{attribute 'pack_mode' := '1'}
TYPE ST_ModulePublishData :
STRUCT
 Header : ST_MqttHeader;
 Devices : ARRAY[0..GVL_PARAM.BAT_MODULE_COUNT-1] OF ST_ModulePublish_V1;
END_STRUCT
END_TYPE

(* stored: Version 1.1.0.1, ProductVersion 3.1.4024.15
   DUT ST_ModulePublishData: Id {19f21c93-ec8a-492d-a3b4-9729765f2a70} *)
